// TIA Portal V21 export
// export: Created 2026-11-10T07:35:21.6795615Z, ExportSetting WithDefaults, DisplayName Totally Integrated Automation Portal, DisplayVersion V21 Update 3, DisplayName STEP 7 Professional, DisplayVersion V21 Update 3, DisplayName STEP 7 Safety, DisplayVersion V21, DisplayName Tech WebApplication, DisplayVersion V21, DisplayName WinCC Basic/Comfort/Advanced, DisplayVersion V21 Update 3, DisplayName WinCC Unified, DisplayVersion V21 Update 3
FUNCTION_BLOCK "FB_Lad_ex148"   // FB72, LAD
{ S7_Optimized_Access := 'TRUE' }
VERSION : 0.1
// stored: AutoNumber true, IsIECCheckEnabled false, IsRetainMemResEnabled false, MemoryReserve 100, SetENOAutomatically false, UDAEnableTagReadback false
   VAR_INPUT
      v_req : Bool;
      v_ret_val : Int;
   END_VAR
   VAR_OUTPUT
      v_busy : Bool;
   END_VAR
   VAR_IN_OUT
      v_srcblk : Variant;
      v_dstblk : Variant;
   END_VAR
BEGIN

REGION Network 1: READ_DBL - Read from data block in the load memory
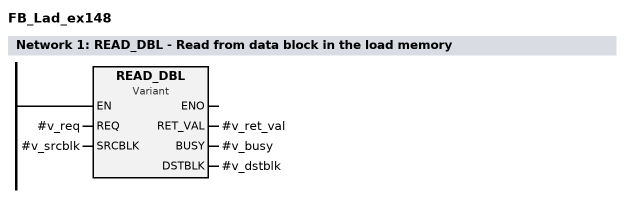
   RUNG wire#powerrail
      { S7_Templates := "[src_type := Variant, dest_type := Variant]" } READ_DBL(REQ := #v_req, SRCBLK := #v_srcblk, RET_VAL => #v_ret_val, BUSY => #v_busy, DSTBLK => #v_dstblk)
   END_RUNG
   // the same network as SCL:
   #v_ret_val := READ_DBL(REQ := #v_req, SRCBLK := #v_srcblk, BUSY => #v_busy, DSTBLK => #v_dstblk);
END_REGION
END_FUNCTION_BLOCK
